// TIA Portal V19 export
DATA_BLOCK "faulty alarms"   // DB20
{ S7_Optimized_Access := 'FALSE'; DB_Accessible_From_OPC_UA := 'FALSE' }
// stored: DBAccessibleFromOPCUA false
   VAR
      faulty_alarms : Struct
         TT01_HIGH : Bool;
         TT02_HIGH : Bool;
         APT01_HIGH : Bool;
         GPT01_HIGH : Bool;
         GPT02_HIGH : Bool;
         GPT03_HIGH : Bool;
         GPT04_HIGH : Bool;
         O2_HIGH : Bool;
         LEL01_HIGH : Bool;
         LEL02_HIGH : Bool;
         PS01_HIGH : Bool;
         TT01_LOW : Bool;
         TT02_LOW : Bool;
         APT01_LOW : Bool;
         GPT01_LOW : Bool;
         GPT02_LOW : Bool;
         GPT03_LOW : Bool;
         GPT04_LOW : Bool;
         O2_LOW : Bool;
         LEL01_LOW : Bool;
         LEL02_LOW : Bool;
         PS01_LOW : Bool;
         TT01_FAULTY : Bool;
         TT02_FAULTY : Bool;
         APT01_FAULTY : Bool;
         GPT01_FAULTY : Bool;
         GPT02_FAULTY : Bool;
         GPT03_FAULTY : Bool;
         GPT04_FAULTY : Bool;
         O2_FAULTY : Bool;
         LEL01_FAULTY : Bool;
         LEL02_FAULTY : Bool;
         PS01_FAULTY : Bool;
         RLT_HIGH : Bool;
         RLT_LOW : Bool;
      END_STRUCT;
   END_VAR
BEGIN
END_DATA_BLOCK
